Fanuc KAREL source: kd00059.KL

-- PROVISIONAL review KL for V1013-1; original PC SHA256 e3750c5f0cf95979e09ff8524cd79bec5109da580b7f392596abbbc36ecb3364
-- Incomplete behavior may be omitted. Consult companion uncertainty JSON. Do not deploy.
PROGRAM KD00059
%NOLOCKGROUP
VAR
  I : INTEGER
  J : INTEGER
  B : BOOLEAN
  R : REAL
  S : STRING[80]
BEGIN
  -- UNRESOLVED_PC offsets 5-18; opcodes 9D,81,18,9D,1B,9D,12,9C,13,04
  -- UNRESOLVED_PC offsets 23-27; opcodes 7F
END KD00059
